Staubli VAL3: getAnaIO.pgx

public program getAnaIO(aio x_aIO, num& x_nValue, bool& x_bError)
  local string l_sDesc
  local string l_sPath
begin
  if ioStatus(x_aIO,l_sDesc,l_sPath)>=0
    x_bError=false
    x_nValue=aioGet(x_aIO)
  else
    x_bError=true
  endIf
end
